(* IEC 61131-3 sources: sis-interlock-demo/tests/POUs/Suites/FB_Voting_Test, 31 files *)

(* ---- AnalogHighInclusiveAtLimit.method.decl.st ---- *)
// Верхняя уставка включительна: 49.99 — норма, ровно 50.0 — требование (2oo3, два канала)
METHOD PRIVATE AnalogHighInclusiveAtLimit
VAR
    fbRig : FB_VotingRig;   // стенд
END_VAR

(* ---- AnalogInfInvalid.method.decl.st ---- *)
// +Inf, -Inf и 1.0E31 (больше REAL_SANE_MAX) — недостоверны; три недостоверных при VoteTrip — ForcedTrip
METHOD PRIVATE AnalogInfInvalid
VAR
    fbRig  : FB_VotingRig;      // стенд
    uPlus  : PL.U_RealBits;     // +Inf
    uMinus : PL.U_RealBits;     // -Inf
END_VAR

(* ---- AnalogLowInclusiveAtLimit.method.decl.st ---- *)
// Нижняя уставка включительна: 10.01 — норма, ровно 10.0 — требование
METHOD PRIVATE AnalogLowInclusiveAtLimit
VAR
    fbRig : FB_VotingRig;   // стенд
END_VAR

(* ---- AnalogNaNInvalid.method.decl.st ---- *)
// NaN при флаге достоверности TRUE — канал недостоверен (событие ChannelInvalid), 2oo3 VoteTrip → 1oo2;
// память гистерезиса канала сбрасывается
METHOD PRIVATE AnalogNaNInvalid
VAR
    fbRig : FB_VotingRig;      // стенд
    uBits : PL.U_RealBits;     // значение REAL по битам IEEE 754
    stEv  : ST_SisEvent;       // событие
END_VAR

(* ---- BypassDeniedWithoutPermit.method.decl.st ---- *)
// Без ключа разрешения запрос байпаса — Denied (BypassDenied); ключ при удержанном запросе ничего не меняет
METHOD PRIVATE BypassDeniedWithoutPermit
VAR
    fbRig : FB_VotingRig;   // стенд
END_VAR

(* ---- BypassEventsWithChannel.method.decl.st ---- *)
// События байпаса несут номер причины, номер канала и метку источника времени
METHOD PRIVATE BypassEventsWithChannel
VAR
    fbRig : FB_VotingRig;   // стенд
    stEv  : ST_SisEvent;    // событие
    ltOn  : LTIME;          // момент включения
END_VAR

(* ---- BypassExpiresExactlyAtMax.method.decl.st ---- *)
// Байпас 10 с недостоверного канала 1: на t0 + 9,9 с действует (канал Bypassed), на t0 + 10,0 с —
// Expired и BypassExpired, канал в том же вызове снова голосует (Invalid)
METHOD PRIVATE BypassExpiresExactlyAtMax
VAR
    fbRig : FB_VotingRig;   // стенд
    stEv  : ST_SisEvent;    // событие
END_VAR

(* ---- BypassLimitLowestChannelWins.method.decl.st ---- *)
// Предел одного байпаса, запросы каналов 2 и 3 в одном вызове: канал 2 — Active, канал 3 — Denied;
// Denied держится до снятия запроса, даже когда место освободилось
METHOD PRIVATE BypassLimitLowestChannelWins
VAR
    fbRig : FB_VotingRig;   // стенд
    stEv  : ST_SisEvent;    // событие
END_VAR

(* ---- BypassPermitLostEnds.method.decl.st ---- *)
// Снятие ключа разрешения заканчивает действующий байпас: Denied и BypassOff, канал снова голосует;
// возврат ключа при удержанном запросе байпас не возобновляет
METHOD PRIVATE BypassPermitLostEnds
VAR
    fbRig : FB_VotingRig;   // стенд
    stEv  : ST_SisEvent;    // событие
END_VAR

(* ---- BypassRemainCountsDown.method.decl.st ---- *)
// Остаток байпаса: 10 с при включении, 7 с через 3 с; после снятия запроса — Off и T#0S
METHOD PRIVATE BypassRemainCountsDown
VAR
    fbRig : FB_VotingRig;   // стенд
END_VAR

(* ---- BypassReRequestNeedsRelease.method.decl.st ---- *)
// После истечения байпаса удержанный запрос его не возобновляет (Expired); снять запрос и подать
// снова — новый байпас на полный срок
METHOD PRIVATE BypassReRequestNeedsRelease
VAR
    fbRig : FB_VotingRig;   // стенд
END_VAR

(* ---- BypassZeroTimeDenied.method.decl.st ---- *)
// tBypassMax = T#0S — байпас запрещён: запрос — Denied
METHOD PRIVATE BypassZeroTimeDenied
VAR
    fbRig : FB_VotingRig;   // стенд
END_VAR

(* ---- CfgAi.method.decl.st ---- *)
// Конфигурация аналоговой группы для тестов: уставка 50.0 (High), гистерезис 2.0, рассогласование
// выключено, байпас до 10 с, один байпас (для 1oo1 — ни одного)
METHOD CfgAi : ST_VotingCfg
VAR_INPUT
    eArch   : E_VoteArch;        // схема
    ePolicy : E_DegradePolicy;   // политика
END_VAR
VAR
    stCfg : ST_VotingCfg;        // результат
END_VAR

(* ---- CfgAi.method.impl.st ---- *)
stCfg.eArch := eArch;
stCfg.ePolicy := ePolicy;
stCfg.eInput := E_SisInputKind.Analog;
stCfg.eLimitDir := E_LimitDir.High;
stCfg.rTripLimit_eu := 50.0;
stCfg.rHyst_eu := 2.0;
stCfg.rDiscrepancyMax_eu := 0.0;
stCfg.tDiscrepancyDelay := T#0S;
stCfg.tBypassMax := T#10S;
IF F_VoteArchChannels(eArch := eArch) > 1 THEN
    stCfg.uiMaxBypass := 1;
ELSE
    stCfg.uiMaxBypass := 0;
END_IF
CfgAi := stCfg;

(* ---- CfgCheckDetectsEachRule.method.decl.st ---- *)
// F_VoteCheckCfg: каждое правило таблицы 4.3 даёт свой бит; верная конфигурация — 0
METHOD PRIVATE CfgCheckDetectsEachRule
VAR
    stCfg : ST_VotingCfg;    // проверяемая конфигурация
    uBad  : U_SisEnumInt;    // значение вне перечисления
    uNaN  : PL.U_RealBits;   // NaN
END_VAR

(* ---- CfgDi.method.decl.st ---- *)
// Конфигурация дискретной группы для тестов: норма канала TRUE, байпас до 10 с, один байпас
// (для 1oo1 — ни одного)
METHOD CfgDi : ST_VotingCfg
VAR_INPUT
    eArch   : E_VoteArch;        // схема
    ePolicy : E_DegradePolicy;   // политика
END_VAR
VAR
    stCfg : ST_VotingCfg;        // результат
END_VAR

(* ---- CfgDi.method.impl.st ---- *)
stCfg.eArch := eArch;
stCfg.ePolicy := ePolicy;
stCfg.eInput := E_SisInputKind.Discrete;
stCfg.xDiHealthy := TRUE;
stCfg.tBypassMax := T#10S;
IF F_VoteArchChannels(eArch := eArch) > 1 THEN
    stCfg.uiMaxBypass := 1;
ELSE
    stCfg.uiMaxBypass := 0;
END_IF
CfgDi := stCfg;

(* ---- CfgErrorRemovesBypasses.method.decl.st ---- *)
// Ошибка конфигурации снимает действующий байпас (CfgError, затем BypassOff), группа срабатывает;
// после исправления удержанный запрос даёт новый байпас на полный срок — таймер не «истёк» за время
// ошибки, потому что вызывался со снятым входом
METHOD PRIVATE CfgErrorRemovesBypasses
VAR
    fbRig : FB_VotingRig;   // стенд
END_VAR

(* ---- ChannelValidityEventsOnChange.method.decl.st ---- *)
// События достоверности — только по смене: исправные каналы при первом вызове событий не дают,
// повтор недостоверности не повторяет событие, возврат — ChannelValid
METHOD PRIVATE ChannelValidityEventsOnChange
VAR
    fbRig : FB_VotingRig;   // стенд
    stEv  : ST_SisEvent;    // событие
END_VAR

(* ---- DefaultCfgTripsCfgError.method.decl.st ---- *)
// Конфигурация по умолчанию (схема None): срабатывание, ошибка VOTE_CFG_ARCH, одно событие CfgError
// с номером причины и кодом ошибки; повторный вызов события не повторяет
METHOD PRIVATE DefaultCfgTripsCfgError
VAR
    fbRig : FB_VotingRig;   // стенд
    stEv  : ST_SisEvent;    // событие
END_VAR

(* ---- DegradeAvailableTwoOfThreeAsTwoOfTwo.method.decl.st ---- *)
// DegradeAvailable, один недостоверный канал 2oo3: действующая схема 2oo2 — один канал Demand не
// срабатывает, два — срабатывают
METHOD PRIVATE DegradeAvailableTwoOfThreeAsTwoOfTwo
VAR
    fbRig : FB_VotingRig;   // стенд
END_VAR

(* ---- DiHealthyFalseInvertsDemand.method.decl.st ---- *)
// xDiHealthy = FALSE: норма — FALSE, требование — TRUE (1oo1)
METHOD PRIVATE DiHealthyFalseInvertsDemand
VAR
    fbRig : FB_VotingRig;   // стенд
END_VAR

(* ---- DiscrepancyAfterDelayExactly.method.decl.st ---- *)
// Разброс 1.5 при допуске 1.0 и задержке 5 с: на t0 + 4,9 с тревоги нет, на t0 + 5,0 с — есть,
// событие DiscrepancyOn с разбросом
METHOD PRIVATE DiscrepancyAfterDelayExactly
VAR
    fbRig : FB_VotingRig;   // стенд
    stEv  : ST_SisEvent;    // событие
END_VAR

(* ---- DiscrepancyAtLimitNoAlarm.method.decl.st ---- *)
// Порог рассогласования строгий: разброс ровно 1.0 при допуске 1.0 — тревоги нет, 1.25 — есть
METHOD PRIVATE DiscrepancyAtLimitNoAlarm
VAR
    fbRig : FB_VotingRig;   // стенд
END_VAR

(* ---- DiscrepancyIgnoresBypassedAndInvalid.method.decl.st ---- *)
// В контроле рассогласования — только каналы Normal и Demand: недостоверный и байпасированный каналы
// не участвуют, при одном участнике разброс 0.0
METHOD PRIVATE DiscrepancyIgnoresBypassedAndInvalid
VAR
    fbRig : FB_VotingRig;   // стенд
END_VAR

(* ---- DiscrepancyNoTripImpact.method.decl.st ---- *)
// Рассогласование — диагностика: тревога есть, требования срабатывания нет
METHOD PRIVATE DiscrepancyNoTripImpact
VAR
    fbRig : FB_VotingRig;   // стенд
END_VAR

(* ---- DiscrepancyZeroDisables.method.decl.st ---- *)
// Допуск 0.0 — контроль рассогласования выключен: разброс 0.0, тревоги нет
METHOD PRIVATE DiscrepancyZeroDisables
VAR
    fbRig : FB_VotingRig;   // стенд
END_VAR

(* ---- HysteresisReleasesBeyondBand.method.decl.st ---- *)
// Гистерезис 2.0 у уставки 50.0 (1oo1): требование держится до 48.0 включительно, снимается при
// 47.99; снизу без памяти 49.0 — норма
METHOD PRIVATE HysteresisReleasesBeyondBand
VAR
    fbRig : FB_VotingRig;   // стенд
END_VAR

(* ---- NoTimeSourceUsesSystemTime.method.decl.st ---- *)
// Без источника времени (itfTime = 0) группа работает от встроенного PL.FB_SystemTime: голосует,
// байпас включается с полным остатком
METHOD PRIVATE NoTimeSourceUsesSystemTime
VAR
    fbVote : FB_Voting;      // ФБ без источника времени
    stIn   : ST_VoteIn;      // входы
    stCmd  : ST_VoteCmd;     // запросы байпаса
    stCfg  : ST_VotingCfg;   // конфигурация
END_VAR

(* ---- TimeBackwardsBypassEnds.method.decl.st ---- *)
// «Время назад» во время байпаса (D-19): срок байпаса недостоверен — байпас заканчивается в том же
// вызове (TimeFault, затем BypassExpired), канал возвращается в голосование; новый байпас — только
// после снятия запроса, и он отсчитывается полностью
METHOD PRIVATE TimeBackwardsBypassEnds
VAR
    fbRig : FB_VotingRig;   // стенд
    ltT0  : LTIME;          // момент включения байпаса
    stEv  : ST_SisEvent;    // событие
END_VAR

(* ---- UnusedChannelsIgnored.method.decl.st ---- *)
// Канал 3 у 1oo2 не входит в схему: требование, недостоверность и запрос байпаса не действуют,
// событий нет, состояние NotUsed
METHOD PRIVATE UnusedChannelsIgnored
VAR
    fbRig : FB_VotingRig;   // стенд
END_VAR
